(* IEC 61131-3 sources: OPEN-PLC-VISION-META-AI-HACKATON/vision-plc-agent/specs/start_lamp_arm, 2 files *)

(* ---- main.st ---- *)
(* start_lamp_arm: start latches the red lamp and moves the arm to 90 deg.
   Stop drives all outputs safe (lamp off, arm to 0) within one scan. *)
PROGRAM Main
VAR
    start_btn AT %IX0.0 : BOOL;
    stop_btn AT %IX0.1 : BOOL;
    lamp_red AT %QX0.0 : BOOL;
    arm_angle AT %QW0 : INT;
    start_edge : R_TRIG; (* rising edge of the start button *)
    stop_edge : R_TRIG;  (* rising edge of the stop button *)
    run_latch : SR;      (* set by start, reset by stop *)
END_VAR

    (* Edge-detect both buttons; never act on a level twice. *)
    start_edge(CLK := start_btn);
    stop_edge(CLK := stop_btn);

    (* Latch the run state; stop wins through the reset input. *)
    run_latch(S1 := start_edge.Q, R := stop_edge.Q);

    (* The stop level forces the safe state in the same scan. *)
    lamp_red := run_latch.Q1 AND NOT stop_btn;
    IF stop_btn THEN
        arm_angle := 0;
    ELSIF run_latch.Q1 THEN
        arm_angle := 90;
    ELSE
        arm_angle := 0;
    END_IF;
END_PROGRAM

(* ---- tests.st ---- *)
(* Acceptance tests for start_lamp_arm, mirroring specs/start_lamp_arm.yaml.
   Single-quoted names: STruC++ v0.7.0 rejects the double-quoted form.
   Tests run in file order; each of the first two drives the program to
   a known state first, so they pass whether or not the SETUP instance
   is shared between tests. *)
SETUP
VAR
    prog : Main;
END_VAR
    prog.start_btn := FALSE;
    prog.stop_btn := FALSE;
END_SETUP

TEST 'start latches lamp and moves arm'
    (* clear any latched state, then pulse start for one scan *)
    prog.stop_btn := TRUE;
    prog();
    prog.stop_btn := FALSE;
    prog.start_btn := TRUE;
    prog();
    prog.start_btn := FALSE;
    prog();
    ASSERT_TRUE(prog.lamp_red);
    ASSERT_EQ(prog.arm_angle, 90);
END_TEST

TEST 'stop clears lamp and homes arm'
    (* latch on first *)
    prog.start_btn := TRUE;
    prog();
    prog.start_btn := FALSE;
    prog();
    ASSERT_TRUE(prog.lamp_red);
    (* press stop: safe state within one scan *)
    prog.stop_btn := TRUE;
    prog();
    ASSERT_FALSE(prog.lamp_red);
    ASSERT_EQ(prog.arm_angle, 0);
    (* release stop: outputs stay safe *)
    prog.stop_btn := FALSE;
    prog();
    ASSERT_FALSE(prog.lamp_red);
    ASSERT_EQ(prog.arm_angle, 0);
END_TEST

TEST 'outputs start safe'
    (* no input yet: lamp off, arm home *)
    prog();
    ASSERT_FALSE(prog.lamp_red);
    ASSERT_EQ(prog.arm_angle, 0);
END_TEST
